FUNCTION_BLOCK Actuator2Op (* Composite Function Block Type *)
  (* Standard: 61499-2 *)
  (* Version 1.0.1, 9/20/2023, ApplicationLibDevTeam, Schneider Electric, First Version *)
  PACKAGE Flexbridge.FestoMPS400;
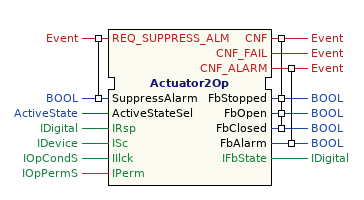
  EVENT_INPUT
    REQ_SUPPRESS_ALM WITH SuppressAlarm; (* Request to update the alarm suppress status *)
  END_EVENT
  EVENT_OUTPUT
    CNF WITH FbOpen, FbClosed, FbStopped; (* Execution confirmation *)
    CNF_FAIL; (* Execution confirmation of failure *)
    CNF_ALARM WITH FbAlarm; (* Execution confirmation of alarm *)
  END_EVENT
  VAR_INPUT
    SuppressAlarm : BOOL; (* 1 = Suppress alarm in HMI *)
    ActiveStateSel : ActiveState; (* Feedback type selection to determine the active state for valves [StateSel configured as Valve1Op or Valve2Op],  0 = Open State  1 = Closed State *)
  END_VAR
  VAR_OUTPUT
    FbStopped : BOOL; (* 1 = Stopped *)
    FbOpen : BOOL; (* 1 = Open *)
    FbClosed : BOOL; (* 1 = Closed *)
    FbAlarm : BOOL; (* 1 = Feedback failure alarm is active *)
  END_VAR
  SOCKETS
    IRsp : IDigital; (* Program remote setpoint interface adapter *)
    ISc : IDevice; (* Sequence control Interface adapter. Controls the block when owner is in program local *)
    IIlck : IOpCondS; (* Interlock condition summary chain input from ilckCondItem blocks *)
    IPerm : IOpPermS; (* Permission condition summary chain input from permCondItem blocks *)
  END_SOCKETS
  PLUGS
    IFbState : IDigital; (* Current feedback status adapter (Value = device feedback status, Status = device alarm data,Bit 1 = Device failure status, Bit 2 = Feedback failure status *)
  END_PLUGS
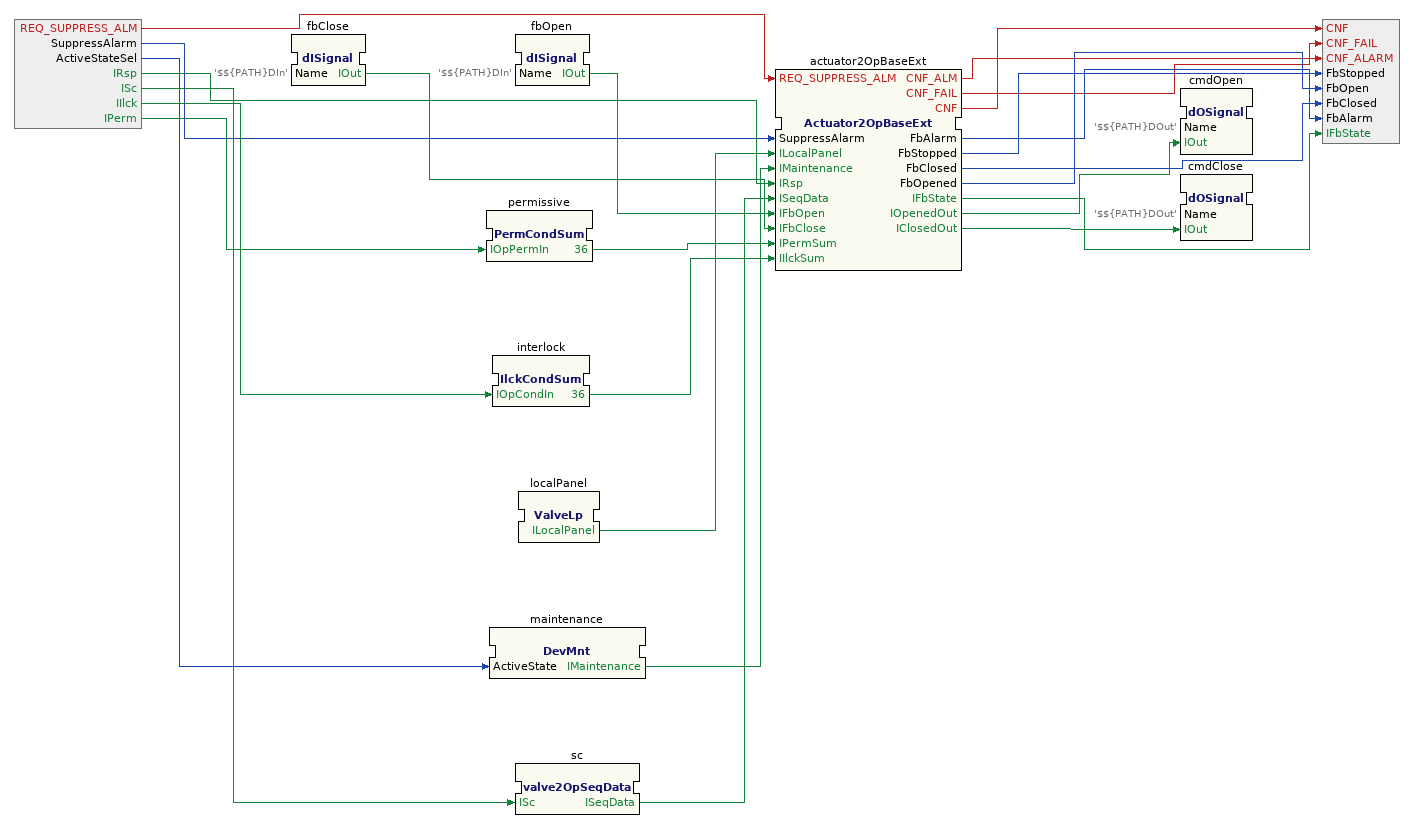
  (* Valve Control *)
  (* Permissive *)
  (* Interlock *)
  (* Sequence Control *)
  (* Local Panel *)
  (* Maintenance *)
  (* Input Hardware Interface *)
  (* Output Hardware Interface *)
  FBS
    interlock : IlckCondSum; {SET_ATTRIBUTE(Configuration.Component.HideUnusedPorts, )}
    permissive : PermCondSum; {SET_ATTRIBUTE(Configuration.Component.HideUnusedPorts, )}
    localPanel : ValveLp; {SET_ATTRIBUTE(Configuration.Component.HideUnusedPorts, )}
    maintenance : DevMnt; {SET_ATTRIBUTE(Configuration.Component.HideUnusedPorts, )}
    sc : valve2OpSeqData;
    fbOpen : dISignal(Name := '$${PATH}DIn'); {SET_ATTRIBUTE(Configuration.Component.HideUnusedPorts, )}
    cmdOpen : dOSignal(Name := '$${PATH}DOut'); {SET_ATTRIBUTE(Configuration.Component.HideUnusedPorts, )}
    fbClose : dISignal(Name := '$${PATH}DIn'); {SET_ATTRIBUTE(Configuration.Component.HideUnusedPorts, )}
    cmdClose : dOSignal(Name := '$${PATH}DOut'); {SET_ATTRIBUTE(Configuration.Component.HideUnusedPorts, )}
    actuator2OpBaseExt : Actuator2OpBaseExt;
  END_FBS
  EVENT_CONNECTIONS
    REQ_SUPPRESS_ALM TO actuator2OpBaseExt.REQ_SUPPRESS_ALM;
    actuator2OpBaseExt.CNF_ALM TO CNF_ALARM;
    actuator2OpBaseExt.CNF_FAIL TO CNF_FAIL;
    actuator2OpBaseExt.CNF TO CNF;
  END_CONNECTIONS
  DATA_CONNECTIONS
    SuppressAlarm TO actuator2OpBaseExt.SuppressAlarm;
    actuator2OpBaseExt.FbAlarm TO FbAlarm;
    actuator2OpBaseExt.FbStopped TO FbStopped;
    actuator2OpBaseExt.FbClosed TO FbClosed;
    actuator2OpBaseExt.FbOpened TO FbOpen;
    ActiveStateSel TO maintenance.ActiveState;
  END_CONNECTIONS
  ADAPTER_CONNECTIONS
    IPerm TO permissive.IOpPermIn;
    ISc TO sc.ISc;
    IIlck TO interlock.IOpCondIn;
    localPanel.ILocalPanel TO actuator2OpBaseExt.ILocalPanel;
    maintenance.IMaintenance TO actuator2OpBaseExt.IMaintenance;
    IRsp TO actuator2OpBaseExt.IRsp;
    sc.ISeqData TO actuator2OpBaseExt.ISeqData;
    actuator2OpBaseExt.IFbState TO IFbState;
    fbOpen.IOut TO actuator2OpBaseExt.IFbOpen;
    fbClose.IOut TO actuator2OpBaseExt.IFbClose;
    permissive.36 TO actuator2OpBaseExt.IPermSum;
    interlock.36 TO actuator2OpBaseExt.IIlckSum;
    actuator2OpBaseExt.IOpenedOut TO cmdOpen.IOut;
    actuator2OpBaseExt.IClosedOut TO cmdClose.IOut;
  END_CONNECTIONS
END_FUNCTION_BLOCK
